Universal Robots URScript: T013_zai-org_GLM-4.7-FP8_baseline_rep1.urscript

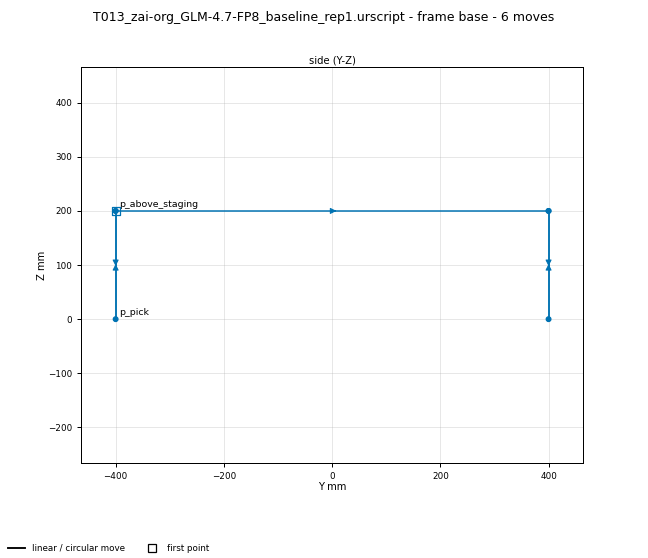
[picture p0: tool path of T013_zai-org_GLM-4.7-FP8_baseline_rep1.urscript in frame base, 6 of 8 moves have a stored position in this frame; points joined in program order, loops and branches not executed]
# UR5e Collaborative Suction Palletizing
# Task: T013 - Light boxes (0.8 kg)
# Mode: Collaborative
# Max TCP Speed: 250.0 mm/s

# --- Configuration ---
# Set TCP (Suction Cup Tool Center Point)
set_tcp(p[0, 0, 0.15, 0, 0, 0])

# Set Payload (Mass in kg, Center of Mass in m)
set_payload(0.8, [0, 0, 0.05])

# --- Waypoint Definitions ---
# Home Position (Joint space)
q_home = [-1.57, -1.57, -1.57, -1.57, -1.57, 0]

# Staging Area (Pick)
p_above_staging = p[0.4, -0.4, 0.2, 2.22, -2.22, 0]
p_pick = p[0.4, -0.4, 0.0, 2.22, -2.22, 0]

# Pallet Area (Place)
p_above_pallet = p[0.4, 0.4, 0.2, 2.22, -2.22, 0]
p_place = p[0.4, 0.4, 0.0, 2.22, -2.22, 0]

# --- Motion Sequence ---

# 1. move_joint: Home, 200.0 mm/s
movej(q_home, a=1.4, v=0.2)

# 2. move_linear: Above staging, 220.0 mm/s
movel(p_above_staging, a=1.2, v=0.22)

# 3. move_linear: Descend to pick, 100.0 mm/s
movel(p_pick, a=0.5, v=0.1)

# Action: Activate Suction
set_digital_out(0, True)
sleep(0.5)

# 4. move_linear: Lift, 180.0 mm/s
movel(p_above_staging, a=1.0, v=0.18)

# 5. move_linear: Transit to pallet, 230.0 mm/s
movel(p_above_pallet, a=1.2, v=0.23)

# 6. move_linear: Descend to place, 100.0 mm/s
movel(p_place, a=0.5, v=0.1)

# Action: Deactivate Suction
set_digital_out(0, False)
sleep(0.5)

# 7. move_linear: Lift from place, 180.0 mm/s
movel(p_above_pallet, a=1.0, v=0.18)

# 8. move_joint: Home, 200.0 mm/s
movej(q_home, a=1.4, v=0.2)

# End of Program
halt
